Yaskawa INFORM job: DEACON.JBI

/JOB
//NAME DEACON
//POS
///NPOS 12,0,0,1,0,0
///TOOL 0
///POSTYPE PULSE
///PULSE
C00000=-203,25202,-52736,-2210,361,1109
C00001=-54,26296,-54047,-3154,2091,1522
C00002=-2459,26373,-53928,20565,2205,-8959
C00003=-1090,24644,-56590,5885,2608,-2440
C00004=-107,26076,-54389,-2560,2158,1257
C00005=-25,22680,-59117,-2562,2858,1234
C00006=-2687,22725,-59051,16788,2967,-7127
C00007=-1476,22541,-59323,8048,2922,-3351
C00008=-1502,21129,-61417,7291,3298,-2989
C00009=-2762,20930,-61711,14924,3436,-6229
C00010=-634,20886,-61775,1677,3337,-588
C00011=-532,16793,-60081,3142,-913,-1276
P00100=0,-60000,-60000,0,-90000,0
//INST
///DATE 2026/06/19 13:14
///ATTR SC,RW
///GROUP1 RB1
NOP
MOVJ P100 VJ=15.00
MOVJ C00000 VJ=15.00
MOVL C00001 V=13.3
ARCON ASF#(13)
MOVC C00002 V=13.3
MOVC C00003 V=13.3
MOVC C00004 V=13.3
ARCOF AEF#(13)
MOVL C00005 V=13.3
ARCON ASF#(13)
MOVL C00006 V=13.3
ARCOF AEF#(13)
MOVL C00007 V=13.3
ARCON ASF#(13)
MOVL C00008 V=13.3
ARCOF AEF#(13)
MOVL C00009 V=13.3
ARCON ASF#(13)
MOVL C00010 V=13.3
ARCOF AEF#(13)
MOVL C00011 V=13.3
MOVJ P100 VJ=15.00
END
